(*
SPDX-FileCopyrightText: © 2026 Oleksandr Tiutyk <trofimich@gmail.com>
SPDX-License-Identifier: MIT
License: https://opensource.org/license/mit
*)

(*!
<summary>Evaluates a branching condition on start and executes either TrueActivity or FalseActivity.</summary>
<description>
Condition is required; TrueActivity and FalseActivity are optional. Selecting a null branch completes
immediately. Resetting resets any non-ready branch activity back to PASSIVE_READY and clears CurrentActivity.
</description>
*)

{attribute 'no_explicit_call' := 'do not call this function block directly'}
{attribute 'enable_dynamic_creation'}
FUNCTION_BLOCK IfElseActivity EXTENDS ExclusiveCompositeActivity
	IMPLEMENTS IIfElseActivity, TOF_Core.IConfigurationSerializable
VAR_STAT
	{attribute 'hide'}
	_ClassName : STRING := __POUNAME();
END_VAR
VAR
	{attribute 'OPC.UA.DA' := '0'}
	_Condition : ICondition;	

	{attribute 'OPC.UA.DA' := '0'}
	_TrueActivity : IActivity;
	
	{attribute 'OPC.UA.DA' := '0'}
	_FalseActivity : IActivity;

	{attribute 'OPC.UA.DA' := '0'}
	_CurrentActivity : IActivity;
END_VAR

(*!
<summary>Borrows the initialized class name used in diagnostics.</summary>
<description>
Returns initialized metadata storage without allocation. Callers must not modify the returned string.
Derived function blocks must use distinct initialized static storage when overriding this metadata.
</description>
*)
{attribute 'monitoring' := 'call'}
PROPERTY ClassName : REFERENCE TO STRING
GET
ClassName REF= _ClassName;
END_GET
END_PROPERTY

(*!
<summary>Returns the branching condition configured for this activity.</summary>
*)
{attribute 'monitoring' := 'call'}
PROPERTY FINAL Condition : ICondition
GET
Condition := _Condition;
END_GET
END_PROPERTY

(*!
<summary>Configures the required branching condition and optional true/false branch activities.</summary>
<description>
Permitted only in PASSIVE_READY. Validates all supplied references before mutating state.
The parent chain and owning workflow must be PASSIVE_READY; fixed workflow association is checked before
mutation. Reusing the same dependency is permitted. Replaced dependencies retain their existing parent links
and must not be attached elsewhere. Parent callbacks are not transactional. Dependencies remain borrowed.
</description>
<param name="condition">Required branching condition.</param>
<param name="trueActivity">Optional activity executed when condition is TRUE.</param>
<param name="falseActivity">Optional activity executed when condition is FALSE.</param>
*)
METHOD Configure
VAR_INPUT
	condition : ICondition; 
	trueActivity : IActivity;
	falseActivity : IActivity;
END_VAR
VAR
END_VAR
IF condition = 0 THEN
	TOF_Core.Exceptions.ThrowArgumentNotSpecified(
		sourceNamespaceName := NamespaceName,
		sourceClassName := ClassName,
		sourcePOUName := __POUNAME(),
		sourcePosition := __POSITION(),
		argumentName := 'condition'
	);
END_IF

IF State <> WORKFLOW_ELEMENT_STATE.PASSIVE_READY THEN
	WorkflowExceptions.ThrowWorkflowConfiguration(
		sourceNamespaceName := NamespaceName,
		sourceClassName := ClassName,
		sourcePOUName := __POUNAME(),
		sourcePosition := __POSITION(),
		message := "Cannot configure IfElseActivity outside PASSIVE_READY"
	);
END_IF

Workflows.ValidateElementAttachment(parent := THIS^, child := condition);

IF trueActivity <> 0 THEN
	ValidateChildActivityAttachment(childActivity := trueActivity, argumentName := 'trueActivity');
END_IF

IF falseActivity <> 0 THEN
	ValidateChildActivityAttachment(childActivity := falseActivity, argumentName := 'falseActivity');
END_IF

IF trueActivity <> 0 AND_THEN trueActivity = falseActivity THEN
	WorkflowExceptions.ThrowWorkflowConfiguration(
		sourceNamespaceName := NamespaceName,
		sourceClassName := ClassName,
		sourcePOUName := __POUNAME(),
		sourcePosition := __POSITION(),
		message := "TrueActivity and FalseActivity cannot reference the same activity instance"
	);
END_IF

_Condition := condition;
_Condition.ParentActivity := THIS^;

_TrueActivity := trueActivity;

IF _TrueActivity <> 0 THEN
	_TrueActivity.ParentActivity := THIS^;
END_IF

_FalseActivity := falseActivity;

IF _FalseActivity <> 0 THEN
	_FalseActivity.ParentActivity := THIS^;
END_IF
END_METHOD

(*!
<summary>Returns the currently selected branch activity, or 0 when none is selected.</summary>
*)
{attribute 'monitoring' := 'call'}
PROPERTY FINAL CurrentActivity : IActivity
GET
CurrentActivity := _CurrentActivity;
END_GET
END_PROPERTY

(*!
<summary>Returns the optional branch activity executed when Condition evaluates to FALSE.</summary>
*)
{attribute 'monitoring' := 'call'}
PROPERTY FINAL FalseActivity : IActivity
GET
FalseActivity := _FalseActivity;
END_GET
END_PROPERTY

(*!
<summary>Borrows the compiler-initialized library namespace.</summary>
<description>
Borrows storage from the live internal namespace provider. Reacquire references after application
reinitialization or relocation. Treat the reference as read-only; no ownership or synchronization is provided.
</description>
*)
{attribute 'monitoring' := 'call'}
PROPERTY NamespaceName : REFERENCE TO STRING
GET
NamespaceName REF= CurrentNamespace.Name;
END_GET
END_PROPERTY

(*!
<summary>Resets any non-ready branch activity back to PASSIVE_READY and clears CurrentActivity.</summary>
<param name="startResetting">TRUE on the initial call from RequestReset.</param>
*)
METHOD PROTECTED OnResetting : ACTIVITY_RESETTING_STATE
VAR_INPUT
	startResetting : BOOL;
END_VAR
IF _TrueActivity <> 0 AND_THEN _TrueActivity.State <> WORKFLOW_ELEMENT_STATE.PASSIVE_READY THEN
	IF ResetChildActivity(childActivity := _TrueActivity) = ACTIVITY_RESETTING_STATE.WORK_IN_PROGRESS THEN
		OnResetting := ACTIVITY_RESETTING_STATE.WORK_IN_PROGRESS;
		RETURN;
	END_IF
END_IF

IF _FalseActivity <> 0 AND_THEN _FalseActivity.State <> WORKFLOW_ELEMENT_STATE.PASSIVE_READY THEN
	IF ResetChildActivity(childActivity := _FalseActivity) = ACTIVITY_RESETTING_STATE.WORK_IN_PROGRESS THEN
		OnResetting := ACTIVITY_RESETTING_STATE.WORK_IN_PROGRESS;
		RETURN;
	END_IF
END_IF

_CurrentActivity := 0;
OnResetting := ACTIVITY_RESETTING_STATE.WORK_RESET;
END_METHOD

(*!
<summary>Evaluates Condition on start to select a branch and advances the selected branch activity.</summary>
<param name="startRunning">TRUE on the initial call of a fresh start.</param>
<param name="startResuming">TRUE on the initial call when resuming from suspension.</param>
<param name="haltReason">Receives the selected branch's HaltReason when halted.</param>
*)
METHOD PROTECTED OnRunning : ACTIVITY_RUNNING_STATE
VAR_INPUT
	startRunning : BOOL;
	startResuming : BOOL;
END_VAR
VAR_OUTPUT
	haltReason : WSTRING(255);
END_VAR
VAR
END_VAR
IF _Condition = 0 THEN
	TOF_Core.Exceptions.ThrowNullReference(
		sourceNamespaceName := NamespaceName,
		sourceClassName := ClassName,
		sourcePOUName := __POUNAME(),
		sourcePosition := __POSITION(),
		variableOrPropertyName := 'Condition'
	);
END_IF

IF startRunning OR_ELSE (startResuming AND_THEN _CurrentActivity = 0) THEN
	IF _Condition.Evaluate(activity := THIS^) THEN
		_CurrentActivity := _TrueActivity;
	ELSE
		_CurrentActivity := _FalseActivity;
	END_IF
END_IF

IF _CurrentActivity <> 0 THEN
	IF startRunning OR_ELSE startResuming THEN
		_CurrentActivity.RequestStart();
	ELSE
		_CurrentActivity.Execute();
	END_IF

	OnRunning := MapChildRunningState(childState := _CurrentActivity.State);

	IF OnRunning = ACTIVITY_RUNNING_STATE.WORK_HALTED THEN
		haltReason := _CurrentActivity.HaltReason;
	END_IF
ELSE
	OnRunning := ACTIVITY_RUNNING_STATE.WORK_COMPLETED;
END_IF
END_METHOD

(*!
<summary>Stops the currently selected branch activity on cancel or suspend.</summary>
<param name="startCancelling">TRUE on the initial call from RequestCancel.</param>
<param name="startSuspending">TRUE on the initial call from RequestSuspend.</param>
<param name="haltReason">Receives the selected branch's HaltReason if it halts while stopping.</param>
*)
METHOD PROTECTED OnStopping : ACTIVITY_STOPPING_STATE
VAR_INPUT
	startCancelling : BOOL;
	startSuspending : BOOL;
END_VAR
VAR_OUTPUT
	haltReason : WSTRING(255);
END_VAR
IF _CurrentActivity = 0 THEN
	OnStopping := ACTIVITY_STOPPING_STATE.WORK_STOPPED;
	RETURN;
END_IF

IF NOT _CurrentActivity.Busy THEN
	IF startCancelling AND_THEN _CurrentActivity.State = WORKFLOW_ELEMENT_STATE.PASSIVE_SUSPENDED THEN
		_CurrentActivity.RequestCancel(reason := _CancelReason);
	END_IF

	OnStopping := MapChildStoppingState(childState := _CurrentActivity.State);

	IF OnStopping = ACTIVITY_STOPPING_STATE.WORK_HALTED THEN
		haltReason := _CurrentActivity.HaltReason;
	END_IF

	RETURN;
END_IF

IF startCancelling THEN
	_CurrentActivity.RequestCancel(reason := _CancelReason);
ELSIF startSuspending THEN
	_CurrentActivity.RequestSuspend();
ELSE
	_CurrentActivity.Execute();
END_IF

OnStopping := MapChildStoppingState(childState := _CurrentActivity.State);

IF OnStopping = ACTIVITY_STOPPING_STATE.WORK_HALTED THEN
	haltReason := _CurrentActivity.HaltReason;
END_IF
END_METHOD

(*!
<summary>Reports the size of this concrete function block instance in bytes.</summary>
<description>
Reports the instance layout rather than dynamic allocations owned by its fields. A derived function block
with a different layout must override this property; the value does not grant disposal rights.
</description>
*)
{attribute 'monitoring' := 'call'}
PROPERTY SelfSize : ULINT
GET
SelfSize := XSIZEOF(THIS^);
END_GET
END_PROPERTY

(*!
<summary>Returns the optional branch activity executed when Condition evaluates to TRUE.</summary>
*)
{attribute 'monitoring' := 'call'}
PROPERTY FINAL TrueActivity : IActivity
GET
TrueActivity := _TrueActivity;
END_GET
END_PROPERTY

(*!
<summary>Writes the configuration fields for this object.</summary>
<description>Borrows the writer for this call. A failure invalidates the current output document.</description>
*)
METHOD Serialize
VAR_INPUT
	writer : TOF_Core.IConfigurationWriter;
END_VAR
Workflows.WriteConfigurationHeader(writer := writer, source := THIS^, displayName := Name, scope := THIS^);
Workflows.WriteConfigurationObject(writer := writer, name := 'condition', source := _Condition);

IF _TrueActivity <> 0 THEN
	Workflows.WriteConfigurationObject(writer := writer, name := 'trueActivity', source := _TrueActivity);
END_IF

IF _FalseActivity <> 0 THEN
	Workflows.WriteConfigurationObject(writer := writer, name := 'falseActivity', source := _FalseActivity);
END_IF
END_METHOD

(*!
<summary>Restores this fresh instance from its configuration object.</summary>
<description>
The reader, document node and deserialization context are borrowed for this call.
On failure discard the partial instance.
</description>
<param name="reader">Active configuration reader.</param>
<param name="node">Configuration node for this activity.</param>
<param name="context">Active configuration deserialization context providing workflow reconstruction services.</param>
*)
METHOD Deserialize
VAR_INPUT
	reader : TOF_Core.IConfigurationReader;
	node : TOF_Core.CONFIGURATION_NODE;
	context : TOF_Core.IConfigurationDeserializationContext;
END_VAR
VAR
	loader : IWorkflowLoader;
END_VAR
loader := WorkflowConfigurationSerializer.ResolveWorkflowLoader(context := context);
Workflows.ReadConfigurationHeader(reader := reader, node := node, target := THIS^, scope := THIS^);

Configure(
	condition := Workflows.ReadCondition(loader := loader, node := reader.GetField(node := node, name := 'condition')),
	trueActivity := Workflows.ReadActivity(loader := loader, node := reader.FindField(node := node, name := 'trueActivity')),
	falseActivity := Workflows.ReadActivity(loader := loader, node := reader.FindField(node := node, name := 'falseActivity'))
);
END_METHOD

END_FUNCTION_BLOCK

(* stored: Version 1.1.0.1
   POU IfElseActivity: Id {1cd30e3c-846b-4eb9-a9ce-7fa6e666beef}, SpecialFunc None
   Folder Overriden methods: Id {7c18294a-5f01-447a-ba92-b48197de5012}
   Property ClassName: Id {6559a5c1-c484-4f35-98d7-b53ed26607c4}
   Get Get: Id {b5af902f-0236-4bda-a28c-5484c06449c6}
   Property Condition: Id {b1a702af-bbd2-41d2-be9e-afd2daed47d9}
   Get Get: Id {f0c499e6-6e86-4678-858a-b550bf5e4979}
   Method Configure: Id {6f8a03c5-4e89-47fe-8a2e-84d291f92130}
   Property CurrentActivity: Id {caf7e17b-b2e7-4778-ae87-9d0c6526b5a9}
   Get Get: Id {536fec86-ac4f-456b-b1d7-f39b6e0344e6}
   Property FalseActivity: Id {38914bcd-273b-46e7-ba69-f901c8bb24c8}
   Get Get: Id {194e2671-2144-4972-955b-4877d38aed87}
   Property NamespaceName: Id {debfe04e-1e73-43a8-995c-aeec5341d752}
   Get Get: Id {b13e4067-e4c9-4850-a82b-05027c911302}
   Method OnResetting: Id {27a480a7-379a-4989-99b6-13fb28dc8329}
   Method OnRunning: Id {f4476714-3be4-4911-b532-89d30e8187a3}
   Method OnStopping: Id {1cb4bb99-ed5f-452b-8916-d1301610d977}
   Property SelfSize: Id {d99b041f-06da-431d-b026-49be93679871}
   Get Get: Id {f7f4d070-b591-40cf-9ba2-fbbac6566838}
   Property TrueActivity: Id {f3b9527e-da8a-43c8-bf8f-24c1c8bff026}
   Get Get: Id {0af70087-f3de-4a61-833c-bfcdd754f1e4}
   Method Serialize: Id {d03455d8-efb5-47b2-ba28-b4a0494cabcf}
   Method Deserialize: Id {db6353eb-6e43-45b5-bf23-80428462a2b0} *)
